// TIA Portal V19 export
FUNCTION_BLOCK "START"   // FB29, LAD
{ S7_Optimized_Access := 'TRUE' }
// stored: MemoryReserve 100, SetENOAutomatically false
   VAR_INPUT
      RUNNING : Bool;
   END_VAR
   VAR_OUTPUT
      START_CMD : Bool;
      STOP_CMD : Bool;
   END_VAR
   VAR_IN_OUT
      "START/STOP" : Bool;
   END_VAR
   VAR
      START_PLS : Bool;
      IEC_Timer_0_Instance { S7_SetPoint := 'True'} : TOF_TIME;
      STOP_PLS : Bool;
      IEC_Timer_0_Instance_1 { S7_SetPoint := 'True'} : TOF_TIME;
      RUNNING_PLS : Bool;
   END_VAR
   VAR_TEMP   // added for the SCL form of the ladder/FBD networks
      _w1 : Bool;
      _w2 : Bool;
      _w3 : Bool;
      _w4 : Bool;
      _w5 : Bool;
   END_VAR
BEGIN

REGION Network 1
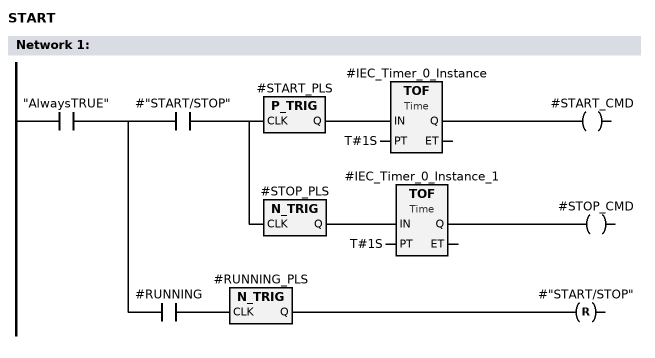
   RUNG wire#powerrail
      Contact( "AlwaysTRUE" )
      wire#w1
      Contact( #"START/STOP" )
      wire#w2
      P_Trig( #START_PLS )
      { S7_Templates := "time_type := Time" } #IEC_Timer_0_Instance.TOF(pt := T#1S, et =>)
      Coil( #START_CMD )
   END_RUNG
   RUNG wire#w2
      N_Trig( #STOP_PLS )
      { S7_Templates := "time_type := Time" } #IEC_Timer_0_Instance_1.TOF(pt := T#1S, et =>)
      Coil( #STOP_CMD )
   END_RUNG
   RUNG wire#w1
      Contact( #RUNNING )
      N_Trig( #RUNNING_PLS )
      R_Coil( #"START/STOP" )
   END_RUNG
   // the same network as SCL:
   #_w1 := "AlwaysTRUE" AND #"START/STOP";
   #_w2 := #_w1 AND NOT #START_PLS;   // rising edge
   #START_PLS := #_w1;
   #IEC_Timer_0_Instance(IN := #_w2, PT := T#1S);   // TOF
   #START_CMD := #IEC_Timer_0_Instance.Q;
   #_w3 := NOT #_w1 AND #STOP_PLS;   // falling edge
   #STOP_PLS := #_w1;
   #IEC_Timer_0_Instance_1(IN := #_w3, PT := T#1S);   // TOF
   #STOP_CMD := #IEC_Timer_0_Instance_1.Q;
   #_w4 := "AlwaysTRUE" AND #RUNNING;
   #_w5 := NOT #_w4 AND #RUNNING_PLS;   // falling edge
   #RUNNING_PLS := #_w4;
   IF #_w5 THEN #"START/STOP" := FALSE; END_IF;
END_REGION
END_FUNCTION_BLOCK
